FUNCTION_BLOCK Prensa_Vibropac (* Prensa desaguadora Vibropac C-Press (VSD-1200) - HidrycoLib *)
  (* Standard: 61499-2 *)
  (* Version 1.1, 12/11/2026, Hidryco, Hidryco, 1.1: modo manual/automatico persistente (LOAD_PERS_DATA no fim da inicializacao). 1.0: Prensa desaguadora Vibropac C-Press (VSD-1200) - tabela Modbus TCP Inovaisa (PV-35525). Campo por symlink ${PATH}: leitura mbR4005..mbR4016 (INT, nome = mbR + registro), mbConexao (connStatusInt, 1 = online); escrita mbW4001 (ciclo remoto 0/1) e mbW4002 (reset 0/1). cfgHabilitada = FALSE para equipamento futuro. *)
  PACKAGE Hidryco.HidrycoLib;
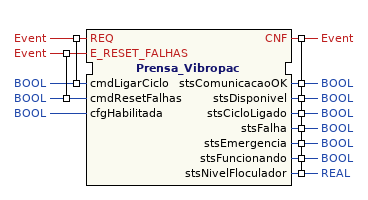
  EVENT_INPUT
    REQ WITH cmdLigarCiclo; (* Atualizacao do processo *)
    E_RESET_FALHAS WITH cmdResetFalhas; (* Reset pelo processo (com cmdResetFalhas = TRUE) *)
  END_EVENT
  EVENT_OUTPUT
    CNF WITH stsComunicacaoOK, stsDisponivel, stsCicloLigado, stsFalha, stsEmergencia, stsFuncionando, stsNivelFloculador; (* Status *)
  END_EVENT
  VAR_INPUT
    cmdLigarCiclo : BOOL; (* TRUE = liga o ciclo remoto do skid (automatico) *)
    cmdResetFalhas : BOOL; (* TRUE = reset (com o evento E_RESET_FALHAS) *)
    cfgHabilitada : BOOL := TRUE; (* FALSE = instancia desabilitada (equipamento futuro) *)
  END_VAR
  VAR_OUTPUT
    stsComunicacaoOK : BOOL; (* Comunicacao Modbus com o CLP do skid OK *)
    stsDisponivel : BOOL; (* Pode ser ligado pelo automatico agora *)
    stsCicloLigado : BOOL; (* Comando de ciclo remoto ligado (4001 = 1) *)
    stsFalha : BOOL; (* Skid em falha (alarme, emergencia ou motor) *)
    stsEmergencia : BOOL; (* Botao de emergencia do skid acionado (4006) *)
    stsFuncionando : BOOL; (* Prensa M1 funcionando *)
    stsNivelFloculador : REAL; (* Nivel do tanque floculador LT1 (%) (4016, 0-1000) *)
  END_VAR
  FBS
    IThis : Prensa_Vibropac_HMI(QI := TRUE);
    plcStart1 : plcStart(Prio := 10);
    Leitura : SYMLINKMULTIVARDST_182274139AA51730B(QI := TRUE, NAME1 := '$${PATH}mbR4005', NAME2 := '$${PATH}mbR4006', NAME3 := '$${PATH}mbR4007', NAME4 := '$${PATH}mbR4008', NAME5 := '$${PATH}mbR4009', NAME6 := '$${PATH}mbR4010', NAME7 := '$${PATH}mbR4011', NAME8 := '$${PATH}mbR4012', NAME9 := '$${PATH}mbR4013', NAME10 := '$${PATH}mbR4014', NAME11 := '$${PATH}mbR4015', NAME12 := '$${PATH}mbR4016'); {SET_ATTRIBUTE(Configuration.GenericFBType.InterfaceParams, Runtime.System#I:=12;VALUE${I$}:INT,INT,INT,INT,INT,INT,INT,INT,INT,INT,INT,INT)}
    Conexao : SYMLINKMULTIVARDST_5A03F112CD5D470(QI := TRUE, NAME1 := '$${PATH}mbConexao'); {SET_ATTRIBUTE(Configuration.GenericFBType.InterfaceParams, Runtime.System#I:=1;VALUE${I$}:INT)}
    EscritaCiclo : SYMLINKMULTIVARSRC_5A03F112CD5D470(QI := TRUE, NAME1 := '$${PATH}mbW4001'); {SET_ATTRIBUTE(Configuration.GenericFBType.InterfaceParams, Runtime.System#I:=1;VALUE${I$}:INT)}
    EscritaReset : SYMLINKMULTIVARSRC_5A03F112CD5D470(QI := TRUE, NAME1 := '$${PATH}mbW4002'); {SET_ATTRIBUTE(Configuration.GenericFBType.InterfaceParams, Runtime.System#I:=1;VALUE${I$}:INT)}
    Logica : basicPrensaVibropac;
    Tick : E_CYCLE(DT := T#1s);
    AlarmeComunicacao : ALARM_BIT(TYPE := 1, ACKTYPE_1 := 2, ACTIVE := TRUE); {SET_ATTRIBUTE(HMI.AlarmText, Prensa sem comunicação)} {SET_ATTRIBUTE(HMI.AlarmClass, Warning)}
    AlarmeEmergencia : ALARM_BIT(TYPE := 1, ACKTYPE_1 := 2, ACTIVE := TRUE); {SET_ATTRIBUTE(HMI.AlarmText, Emergência acionada na prensa)}
    AlarmeSkid : ALARM_BIT(TYPE := 1, ACKTYPE_1 := 2, ACTIVE := TRUE); {SET_ATTRIBUTE(HMI.AlarmText, Alarme no painel do skid da prensa)}
    AlarmeMotor : ALARM_BIT(TYPE := 1, ACKTYPE_1 := 2, ACTIVE := TRUE); {SET_ATTRIBUTE(HMI.AlarmText, Falha de motor da prensa)}
  END_FBS
  EVENT_CONNECTIONS
    plcStart1.FIRST_INIT TO IThis.772F361DFDEA6D62;
    plcStart1.REDO_INIT TO IThis.772F361DFDEA6D62;
    IThis.BF94B10C197EACBD TO Leitura.INIT;
    Leitura.INITO TO Conexao.INIT;
    Conexao.INITO TO EscritaCiclo.INIT;
    EscritaCiclo.INITO TO EscritaReset.INIT;
    EscritaReset.INITO TO Logica.D299CD8A82E1136D;
    Logica.8E1980C6681EA422 TO Tick.START;
    Logica.8E1980C6681EA422 TO AlarmeComunicacao.INIT;
    AlarmeComunicacao.INITO TO AlarmeComunicacao.REQ_INITDATA;
    AlarmeComunicacao.CNF_INITDATA TO AlarmeComunicacao.ACTIVATE;
    AlarmeEmergencia.INITO TO AlarmeEmergencia.REQ_INITDATA;
    AlarmeEmergencia.CNF_INITDATA TO AlarmeEmergencia.ACTIVATE;
    AlarmeComunicacao.INITO TO AlarmeEmergencia.INIT;
    AlarmeSkid.INITO TO AlarmeSkid.REQ_INITDATA;
    AlarmeSkid.CNF_INITDATA TO AlarmeSkid.ACTIVATE;
    AlarmeEmergencia.INITO TO AlarmeSkid.INIT;
    AlarmeMotor.INITO TO AlarmeMotor.REQ_INITDATA;
    AlarmeMotor.CNF_INITDATA TO AlarmeMotor.ACTIVATE;
    AlarmeSkid.INITO TO AlarmeMotor.INIT;
    AlarmeMotor.INITO TO plcStart1.ACK_FIRST;
    Leitura.CNF TO Logica.A0D070BFB6922E53;
    Conexao.CNF TO Logica.17E947DFA2FE7501;
    Tick.EO TO Logica.F8A0187FBB813D55;
    REQ TO Logica.06851BFC2F886180;
    E_RESET_FALHAS TO Logica.E47BD40336CF9E69;
    Logica.2C24C509F6C5D681 TO CNF;
    IThis.53010F5E5B460566 TO Logica.626A32EF4848BC0C;
    IThis.2255219503064CD0 TO Logica.83A35AA7A419EBC5;
    IThis.2686D00AC42141DA TO Logica.178824CC6CD635F9;
    Logica.6190852B9B096605 TO IThis.BC72739772237053;
    Logica.6190852B9B096605 TO AlarmeComunicacao.REQ;
    AlarmeComunicacao.IND_1 TO IThis.BC72739772237053;
    IThis.2686D00AC42141DA TO AlarmeComunicacao.ACK_C1;
    E_RESET_FALHAS TO AlarmeComunicacao.ACK_C1;
    Logica.6190852B9B096605 TO AlarmeEmergencia.REQ;
    AlarmeEmergencia.IND_1 TO IThis.BC72739772237053;
    IThis.2686D00AC42141DA TO AlarmeEmergencia.ACK_C1;
    E_RESET_FALHAS TO AlarmeEmergencia.ACK_C1;
    Logica.6190852B9B096605 TO AlarmeSkid.REQ;
    AlarmeSkid.IND_1 TO IThis.BC72739772237053;
    IThis.2686D00AC42141DA TO AlarmeSkid.ACK_C1;
    E_RESET_FALHAS TO AlarmeSkid.ACK_C1;
    Logica.6190852B9B096605 TO AlarmeMotor.REQ;
    AlarmeMotor.IND_1 TO IThis.BC72739772237053;
    IThis.2686D00AC42141DA TO AlarmeMotor.ACK_C1;
    E_RESET_FALHAS TO AlarmeMotor.ACK_C1;
    Logica.1569871310BFDF0C TO EscritaCiclo.REQ;
    Logica.1569871310BFDF0C TO EscritaReset.REQ;
    AlarmeMotor.INITO TO IThis.DFDF002DEBBD14C7;
  END_CONNECTIONS
  DATA_CONNECTIONS
    Leitura.VALUE1 TO Logica.1F794C4FB36A8D3D;
    Leitura.VALUE2 TO Logica.8CADB224D47AF0CD;
    Leitura.VALUE3 TO Logica.5DDE49FF5C910A23;
    Leitura.VALUE4 TO Logica.EF5E189ABE367D0A;
    Leitura.VALUE5 TO Logica.0F7C3839F37D1CA5;
    Leitura.VALUE6 TO Logica.AE64E46748097A8C;
    Leitura.VALUE7 TO Logica.2C3F5F0650E06C3B;
    Leitura.VALUE8 TO Logica.D3DFEC8C186074CF;
    Leitura.VALUE9 TO Logica.43F79E76B893B9EA;
    Leitura.VALUE10 TO Logica.DC4D6BA5F042BA7A;
    Leitura.VALUE11 TO Logica.80C9DBC9EBE9F1D4;
    Leitura.VALUE12 TO Logica.6F2F5BCB899CFD50;
    Conexao.VALUE1 TO Logica.7EEF417EA22477A6;
    cmdLigarCiclo TO Logica.1F60AF7D7A308712;
    cfgHabilitada TO Logica.730469C1CCCA35EA;
    cmdResetFalhas TO Logica.AF09E58A3FCA6901;
    Logica.0EDA92400C074EF2 TO stsComunicacaoOK;
    Logica.D66869E7164BDDA8 TO stsDisponivel;
    Logica.E72A00ED464B6A3E TO stsCicloLigado;
    Logica.D42679A497B20E1C TO stsFalha;
    Logica.6E23A010B6958DC5 TO stsEmergencia;
    Logica.4066B64CEA148923 TO stsFuncionando;
    Logica.031B294E0F64A3F3 TO stsNivelFloculador;
    IThis.F54A43FCFF519AD6 TO Logica.054295709C415D9E;
    IThis.357B0E799A2B2CD7 TO Logica.61BDC569ABCE85FC;
    IThis.8EBA7C7431C58F42 TO Logica.6DC22945A4E84395;
    Logica.0EDA92400C074EF2 TO IThis.2D3631F568A49914;
    Logica.5BAEBAB6BBAFB013 TO IThis.67AD409CE58402E3;
    Logica.078A8C2377AAD51F TO IThis.0648DCCB0DE07BD9;
    Logica.C3C42C252D3065A4 TO IThis.2FAB077B4C5A2AB5;
    Logica.E72A00ED464B6A3E TO IThis.F32DF3573AA446BD;
    Logica.48D39DA57D78D766 TO IThis.BE39F232CA8B869D;
    Logica.32D2B033B0FC9F12 TO IThis.13F85277C82B8A59;
    Logica.6E23A010B6958DC5 TO IThis.0B5961717B048ABD;
    Logica.097B012F90436A1C TO IThis.15A055430FA2F9FC;
    Logica.D42679A497B20E1C TO IThis.A94E40D540FA592B;
    Logica.D66869E7164BDDA8 TO IThis.0FDB015378C04C5D;
    Logica.37D6D5FA2F9DE978 TO IThis.C4A372EB5C510CCB;
    Logica.00910A4964C2ECC0 TO IThis.E66E6AAAE6FC88AC;
    Logica.AFCF91D8E0A45F8A TO IThis.4F0B9502D8E097C4;
    Logica.69561591E596F7A6 TO IThis.9BCF7F1DAE064FD1;
    Logica.4E5C009C6407D637 TO IThis.B815E58E6B24CA97;
    Logica.58E95E51C9C3528D TO IThis.5DA1D9B02B17694E;
    Logica.B1A1392CB5C49FB3 TO IThis.54DF2D1189A782D7;
    Logica.B468D8458D1D2D2D TO IThis.3EE625D397F38686;
    Logica.1B82EB2F2B07282B TO IThis.EB2C13022E0703B0;
    Logica.EF9D7378E302155F TO IThis.47E587401749CA49;
    Logica.031B294E0F64A3F3 TO IThis.CFCBD5C9BB134D43;
    Logica.4066B64CEA148923 TO IThis.7834DDF8B8A67BB9;
    Logica.5BAEBAB6BBAFB013 TO AlarmeComunicacao.INP;
    AlarmeComunicacao.STATE_1 TO IThis.912B7B6248333678;
    Logica.6E23A010B6958DC5 TO AlarmeEmergencia.INP;
    AlarmeEmergencia.STATE_1 TO IThis.B52B8FE2067186A0;
    Logica.32D2B033B0FC9F12 TO AlarmeSkid.INP;
    AlarmeSkid.STATE_1 TO IThis.DAB162B603363F91;
    Logica.097B012F90436A1C TO AlarmeMotor.INP;
    AlarmeMotor.STATE_1 TO IThis.D1F404D2A05AA8AD;
    Logica.61BC6C8F0F362AE8 TO EscritaCiclo.VALUE1;
    Logica.7FDD9720F54034D7 TO EscritaReset.VALUE1;
  END_CONNECTIONS
END_FUNCTION_BLOCK
